(* IEC 61131-3 sources: sis-interlock-demo/src/POUs/Sis/F_SisFirstBit, 2 files *)

(* ---- F_SisFirstBit.decl.st ---- *)
// Назначение: индекс младшего установленного бита маски с единицы (бит 0 — 1); 0 — битов нет.
//             Первопричина и причина события EffectTrip — младший индекс (разделы 6.6, 6.7).
// Автор:      kr0nsch
// Версия:     0.1.0
// Документ:   docs/DESIGN.md, раздел «8.2 Функции работы с битами»
// ВНИМАНИЕ:   код демонстрационный и не предназначен для систем безопасности. Реальная ПАЗ
//             требует определения SIL, сертифицированных аппаратных и программных средств
//             и валидации по ГОСТ Р МЭК 61511.
FUNCTION F_SisFirstBit : UINT
VAR_INPUT
    wMask : WORD;    // маска
END_VAR
VAR
    uiIdx   : UINT;  // проверяемый индекс
    uiFound : UINT;  // найденный индекс; 0 — ещё не найден
END_VAR

(* ---- F_SisFirstBit.impl.st ---- *)
uiFound := 0;
FOR uiIdx := 1 TO GVL_Const.WORD_BITS DO
    IF uiFound = 0 AND F_SisBit(wMask := wMask, uiIdx := uiIdx) THEN
        uiFound := uiIdx;
    END_IF
END_FOR
F_SisFirstBit := uiFound;
